FUNCTION_BLOCK SECOND_ORDER_PROCESS (* Offline identification prototype; see docs/adaptive/4diac-design.md *)
  (* Standard: 61499-2 *)
  (* Version 0.1, 2026-09-26, Guilherme *)
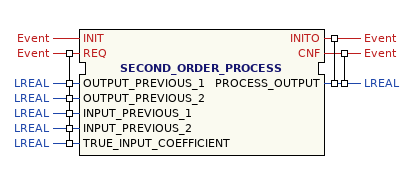
  EVENT_INPUT
    INIT;
    REQ WITH OUTPUT_PREVIOUS_1, OUTPUT_PREVIOUS_2, INPUT_PREVIOUS_1, INPUT_PREVIOUS_2, TRUE_INPUT_COEFFICIENT;
  END_EVENT
  EVENT_OUTPUT
    INITO WITH PROCESS_OUTPUT;
    CNF WITH PROCESS_OUTPUT;
  END_EVENT
  VAR_INPUT
    OUTPUT_PREVIOUS_1 : LREAL;
    OUTPUT_PREVIOUS_2 : LREAL;
    INPUT_PREVIOUS_1 : LREAL;
    INPUT_PREVIOUS_2 : LREAL;
    TRUE_INPUT_COEFFICIENT : LREAL;
  END_VAR
  VAR_OUTPUT
    PROCESS_OUTPUT : LREAL;
  END_VAR
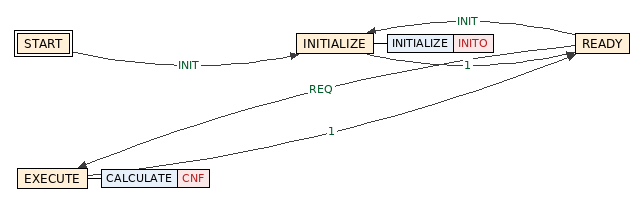
  EC_STATES
    START;
    INITIALIZE : INITIALIZE -> INITO;
    READY;
    EXECUTE : CALCULATE -> CNF;
  END_STATES
  EC_TRANSITIONS
    START TO INITIALIZE := INIT;
    INITIALIZE TO READY := 1;
    READY TO INITIALIZE := INIT;
    READY TO EXECUTE := REQ;
    EXECUTE TO READY := 1;
  END_TRANSITIONS
  ALGORITHM INITIALIZE IN ST:
PROCESS_OUTPUT := 0.0;
  END_ALGORITHM
  ALGORITHM CALCULATE IN ST:
PROCESS_OUTPUT := 1.2 * OUTPUT_PREVIOUS_1 - 0.36 * OUTPUT_PREVIOUS_2 + TRUE_INPUT_COEFFICIENT * INPUT_PREVIOUS_1 + 0.06 * INPUT_PREVIOUS_2;
  END_ALGORITHM
END_FUNCTION_BLOCK
